Fanuc KAREL source: kt00598.KL

-- PROVISIONAL review KL for V1013-1; original PC SHA256 e1b3099f34d9add6a6536116dccecd6314946f22847cded3cd65ddf6d61a26ff
-- Incomplete behavior may be omitted. Consult companion uncertainty JSON. Do not deploy.
PROGRAM KT00598
%NOLOCKGROUP
VAR
  I1 : INTEGER
  I2 : INTEGER
  OUT : INTEGER
BEGIN
  -- UNRESOLVED_PC offsets 5-16; opcodes 2E,23
  -- UNRESOLVED_PC offsets 21-32; opcodes 2E,23
  -- UNRESOLVED_PC offsets 37-48; opcodes 2E,23
  -- UNRESOLVED_PC offsets 53-64; opcodes 2E,23
  -- UNRESOLVED_PC offsets 69-82; opcodes 21,48,23
  -- UNRESOLVED_PC offsets 87-91; opcodes 7F
END KT00598
